(* CODESYS project FeedRobot.xml

Project tree, tasks and I/O mapping:
  visualisation FeedRobot
*)

// /FeedRobot
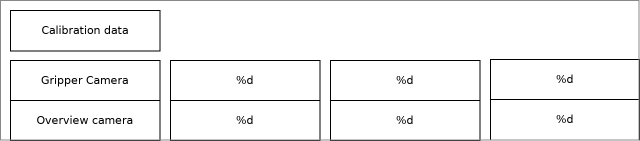
VISUALIZATION FeedRobot  // 640x141
    Rectangle (10,10 150x41), "Calibration data"
    Rectangle (10,60 150x41), "Gripper Camera"
    Rectangle (170,60 150x41), "%d", text variable: PersistentVars.scFeedrobot.CameraGripper.ascCameraCalibration[1].RotationCenter.PosX
    Rectangle (330,60 150x41), "%d", text variable: PersistentVars.scFeedrobot.CameraGripper.ascCameraCalibration[1].RotationCenter.PosY
    Rectangle (10,100 150x41), "Overview camera"
    Rectangle (170,100 150x41), "%d", text variable: PersistentVars.scFeedrobot.CameraAngle.ascCameraCalibration[1].RotationCenter.PosX
    Rectangle (330,100 150x41), "%d", text variable: PersistentVars.scFeedrobot.CameraAngle.ascCameraCalibration[1].RotationCenter.PosY
    Rectangle (490,59 150x41), "%d", text variable: PersistentVars.scFeedrobot.CameraGripper.ascCameraCalibration[1].scale
    Rectangle (490,99 150x41), "%d", text variable: PersistentVars.scFeedrobot.CameraAngle.ascCameraCalibration[1].scale
END_VISUALIZATION
